Fanuc KAREL source: KT00519.KL

PROGRAM KT00519
%NOLOCKGROUP
VAR
  P1: XYZWPREXT
  P2: XYZWPR
  OUT: POSITION
BEGIN
  P1.X = 1.0
    P2.Y = 2.0
  OUT = P1 : P2
END KT00519
